// TIA Portal V19 export
VAR_GLOBAL   // PLC tag table "R2_IN"
   "ByteIN :0 R2" AT %IB218 : Byte;   // System Bits 1
   "ByteIN :1 R2" AT %IB219 : Byte;   // System Bits 2
   "ByteIN :2 R2" AT %IB220 : Byte;   // Signals
   "ByteIN :3 R2" AT %IB221 : Byte;   // Signals
   "ByteIN :4 R2" AT %IB222 : Byte;   // CMD
   "ByteIN :5 R2" AT %IB223 : Byte;
   "ByteIN :6 R2" AT %IB224 : Byte;
   "ByteIN :7 R2" AT %IB225 : Byte;
   "ByteIN :8 R2" AT %IB226 : Byte;
   "ByteIN :9 R2" AT %IB227 : Byte;
   "ByteIN :10 R2" AT %IB228 : Byte;
   "ByteIN :11 R2" AT %IB229 : Byte;
   "ByteIN :12 R2" AT %IB230 : Byte;
   "ByteIN :13 R2" AT %IB231 : Byte;
   "ByteIN :14 R2" AT %IB232 : Byte;
   "ByteIN :15 R2" AT %IB233 : Byte;
   "ByteIN :16 R2" AT %IB234 : Byte;
   "ByteIN :17 R2" AT %IB235 : Byte;
   "ByteIN :18 R2" AT %IB236 : Byte;
   "ByteIN :19 R2" AT %IB237 : Byte;
   "ByteIN :20 R2" AT %IB238 : Byte;
   "ByteIN :21 R2" AT %IB239 : Byte;
   "ByteIN :22 R2" AT %IB240 : Byte;
   "ByteIN :23 R2" AT %IB241 : Byte;
   "ByteIN :24 R2" AT %IB242 : Byte;
   "ByteIN :25 R2" AT %IB243 : Byte;
   "ByteIN :26 R2" AT %IB244 : Byte;
   "ByteIN :27 R2" AT %IB245 : Byte;
   "ByteIN :28 R2" AT %IB246 : Byte;
   "ByteIN :29 R2" AT %IB247 : Byte;
   "ByteIN :30 R2" AT %IB248 : Byte;
   "ByteIN :31 R2" AT %IB249 : Byte;
   "ByteIN :32 R2" AT %IB250 : Byte;
   "ByteIN :33 R2" AT %IB251 : Byte;
   "ByteIN :34 R2" AT %IB252 : Byte;
   "ByteIN :35 R2" AT %IB253 : Byte;
   "ByteIN :36 R2" AT %IB254 : Byte;
   "ByteIN :37 R2" AT %IB255 : Byte;
   "ByteIN :38 R2" AT %IB256 : Byte;
   "ByteIN :39 R2" AT %IB257 : Byte;
   "ByteIN :40 R2" AT %IB258 : Byte;
   "ByteIN :41 R2" AT %IB259 : Byte;
   "ByteIN :42 R2" AT %IB260 : Byte;
   "ByteIN :43 R2" AT %IB261 : Byte;
   "ByteIN :44 R2" AT %IB262 : Byte;
   "ByteIN :45 R2" AT %IB263 : Byte;
   "ByteIN :46 R2" AT %IB264 : Byte;
   "ByteIN :47 R2" AT %IB265 : Byte;
   "ByteIN :48 R2" AT %IB266 : Byte;
   "ByteIN :49 R2" AT %IB267 : Byte;
   "ByteIN :50 R2" AT %IB268 : Byte;
   "ByteIN :51 R2" AT %IB269 : Byte;
   "ByteIN :52 R2" AT %IB270 : Byte;
   "ByteIN :53 R2" AT %IB271 : Byte;
   "ByteIN :54 R2" AT %IB272 : Byte;
   "ByteIN :55 R2" AT %IB273 : Byte;
   "ByteIN :56 R2" AT %IB274 : Byte;
   "ByteIN :57 R2" AT %IB275 : Byte;
   "ByteIN :58 R2" AT %IB276 : Byte;
   "ByteIN :59 R2" AT %IB277 : Byte;
   "ByteIN :60 R2" AT %IB278 : Byte;
   "ByteIN :61 R2" AT %IB279 : Byte;
   "ByteIN :62 R2" AT %IB280 : Byte;
   "ByteIN :63 R2" AT %IB281 : Byte;
END_VAR
